{region 'Documentation'}
(*!
<summary>Check that IN is strictly earlier than Maximum.</summary>
*)
{endregion}
FUNCTION_BLOCK AssertEarlierThan_DT EXTENDS AssertionBase
VAR_INPUT
    IN : DT; //! Actual value checked or observed by this Assertion.
    Maximum : DT; //! Exclusive upper bound; the actual value or count must be smaller.
END_VAR

SUPER^();

{region 'Documentation'}
(*!
<summary>Evaluate the typed temporal relation and report higher-priority errors first.</summary>
*)
{endregion}
METHOD PROTECTED Assert
VAR
    Message : STRING(GVL_Constants.MessageLength);
    MaximumText : STRING(GVL_Constants.AssertionValueLength);
    ActualText : STRING(GVL_Constants.AssertionValueLength);
END_VAR
IF NOT EvaluationActive THEN
    RETURN;
END_IF;

IF Result = E_Result.Error THEN
    RETURN;
END_IF;

IF Result = E_Result.Failed THEN
    RETURN;
END_IF;

IF IN >= Maximum THEN
    MaximumText := DT_TO_STRING(Maximum);
    ActualText := DT_TO_STRING(IN);
    Message := CONCAT('Assertion failed: value is not earlier than limit. Maximum = ',
        MaximumText);
    Message := CONCAT(Message, ', Actual = ');
    Message := CONCAT(Message, ActualText);
    Message := CONCAT(Message, '.');
    Fail(Message := Message);
    RETURN;
END_IF;

Pass();
END_METHOD

END_FUNCTION_BLOCK

(* stored: Version 1.1.0.1
   POU AssertEarlierThan_DT: Id {e98944ad-320b-46ca-a483-0128db4479b9}, SpecialFunc None
   Folder Internal: Id {e0c802f1-b2d7-4cc8-a944-562ca957f26b}
   Method Assert: Id {866aeeb6-fa8e-49b5-b620-7553c76f9023} *)
